(* IEC 61131-3 sources: PLC-Static-Analysis/modules/plc-rules/src/test/resources/PLCA-L021, 2 files *)

(* ---- compliant.st ---- *)
PROGRAM P_L021ok
VAR
    n : INT;
    m : INT;
    r : REAL;
    b : BOOL;
    c : BOOL;
    q : BOOL;
END_VAR
IF n > 10 THEN
    // handled by the alarm task
END_IF
CASE n OF
    1: q := TRUE;
    2: (* idle: wait for start *)
ELSE
    (* unknown step: ignored on purpose *)
END_CASE
IF n > 10 THEN
ELSE
    q := TRUE;
END_IF
END_PROGRAM

(* ---- noncompliant.st ---- *)
PROGRAM P_L021
VAR
    n : INT;
    m : INT;
    r : REAL;
    b : BOOL;
    c : BOOL;
    q : BOOL;
END_VAR
(* PLCA-L021 *) IF n > 10 THEN
END_IF
IF n > 10 THEN
    q := TRUE;
ELSIF (* PLCA-L021 *) n > 5 THEN
ELSE
    q := FALSE;
END_IF
IF n > 10 THEN
    q := TRUE;
(* PLCA-L021 *) ELSE
END_IF
CASE n OF
    1: q := TRUE;
    (* PLCA-L021 *) 2:
END_CASE
CASE n OF
    1: q := TRUE;
(* PLCA-L021 *) ELSE
END_CASE
END_PROGRAM
